TYPE ST_Point2D :
STRUCT
    X : LREAL; // Tọa độ X (mm)
    Y : LREAL; // Tọa độ Y (mm)
END_STRUCT
END_TYPE

(* stored: Version 1.1.0.1, ProductVersion 3.1.4024.16
   DUT ST_Point2D: Id {c4d17d3d-73dd-4963-b025-dcc5a75bd680} *)
